(* IEC 61131-3 sources: tsplc/packages/vscode-extension/tests/fixtures/blueprint/types/ST_Sorter, 3 files *)

(* ---- ST_Sorter.st ---- *)
(*
Zone controls, routing context, and transfer status for a two-zone right-angle sorter.
*)
TYPE ST_Sorter :
STRUCT
	(* Two zone controllers in the sorter assembly; each zone has its own control outputs and feedback. *)
	Zones : ARRAY[1..2] OF ST_MotorZone;
	(* Transfer sequence observations; these are not zone controller registers. *)
	Status : ST_SorterStatus;
	(* PLC-owned routing context, never mapped directly to electrical outputs. *)
	Routing : ST_SorterRouting;
END_STRUCT
END_TYPE

(* ---- ST_SorterRouting.st ---- *)
(*
Zone controls, routing context, and transfer status for a two-zone right-angle sorter.
*)
TYPE ST_SorterRouting :
STRUCT
	(* 0=unknown; 1..4=configured pallet lane. Unknown must hold. *)
	PalletLane : INT;
	(* Identity to which the requested route applies. *)
	CommandPayload : STRING(80);
	(* PlantConstants.Product*: 0=unknown, 1=still, 2=sparkling, 3=juice. *)
	ProductType : INT;
	(* Payload is a crate with no remaining bottles. *)
	EmptyCrate : BOOL;
	(* Payload requires inspection before release. *)
	NeedsInspection : BOOL;
	(* Derived from receiving sensors, enable state, and reservations; not a reader observation. *)
	ReceivingAvailable : BOOL;
	(* Assigned station identity. Direction is resolved by configured port mapping. *)
	TargetStation : STRING(80);
END_STRUCT
END_TYPE

(* ---- ST_SorterStatus.st ---- *)
(*
Zone controls, routing context, and transfer status for a two-zone right-angle sorter.
*)
TYPE ST_SorterStatus :
STRUCT
	(* FALSE until the owning PLC logic supplies a current status; FALSE on stale or unavailable inputs. *)
	Valid : BOOL;
	(* Committed transfer route, not a measured actuator position. PlantConstants.Route*: 0=none/hold, 1=through, 2=left, 3=right. Logical ports; no actuator wiring implied. *)
	ActiveRoute : INT;
	(* Transfer is in progress until configured arrival feedback completes it. *)
	Busy : BOOL;
	(* Fault in the actuator interface or transfer sequence. *)
	Faulted : BOOL;
	(* Payload currently committed to a transfer; cleared once arrival is confirmed. *)
	TransferPayload : STRING(80);
END_STRUCT
END_TYPE
